Fanuc KAREL source: KT00501.KL

PROGRAM KT00501
%NOLOCKGROUP
VAR
  P1: XYZWPR
  P2: XYZWPR
  OUT: XYZWPREXT
BEGIN
  P1.X = 1.0
  P2.Y = 2.0
  P1.X = 1.0
  P2.Y = 2.0
  OUT = P1 : P2
END KT00501
